Fanuc KAREL source: kt00165.KL

-- PROVISIONAL review KL for V940-1; original PC SHA256 c3caafa371b7edd64d8483402ecccb006a0d35ddf0b30ee1f7e7dd5537d50c46
-- Incomplete behavior may be omitted. Consult companion uncertainty JSON. Do not deploy.
PROGRAM KT00165
%NOLOCKGROUP
VAR
  I1 : INTEGER
  OUT : INTEGER
-- UNRESOLVED_DECL Y2 type=002018
BEGIN
  -- V9_ZERO_TABLE_METADATA_HINT layout=0001; no indexed target words; source/name/runtime held
  -- UNRESOLVED_PC offsets 5-16; opcodes 2E,23
  -- UNRESOLVED_PC offsets 21-35; opcodes 2E,22,9D,33,B2
  -- UNRESOLVED_PC offsets 40-62; opcodes 21,22,9D,33,B1,56,23
  -- UNRESOLVED_PC offsets 67-71; opcodes 7F
END KT00165
